FUNCTION_BLOCK UCT_PreTratamento_HMI (* Service Interface Function Block Type *)
  (* Standard: 61499-2 *)
  (* Version 1.5, 04/11/2026, Hidryco, Hidryco, 1.5: STS_LIGADO, STS_AUTOMATICO (IO List da Nereda). IHM da UCT (nomes do IThis do Pre_Tratamento antigo) *)
  PACKAGE Hidryco.HidrycoLib;
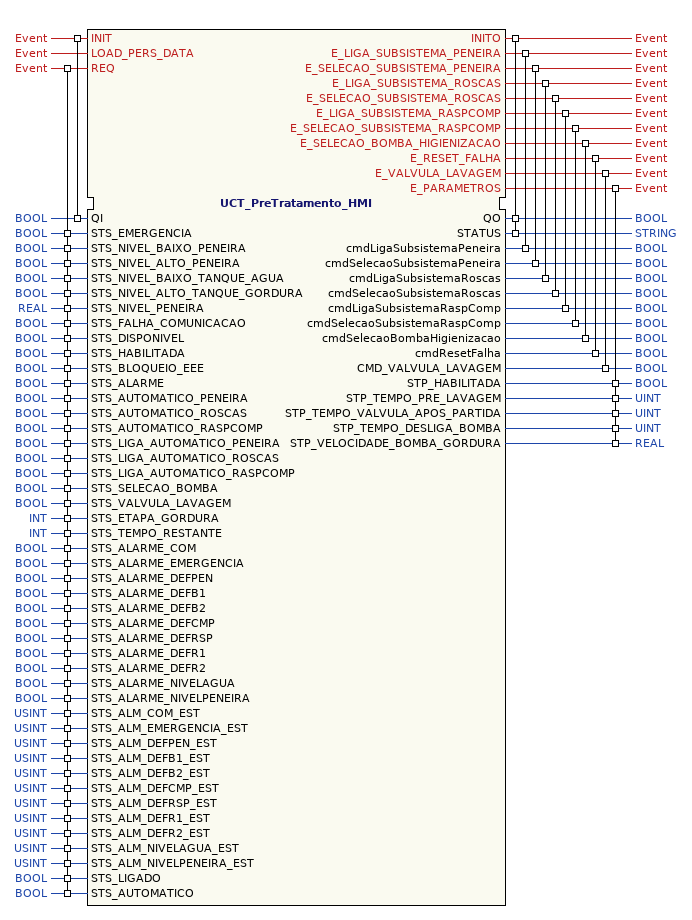
  EVENT_INPUT
    INIT WITH QI;
    LOAD_PERS_DATA; (* Reenvia os parametros persistentes *)
    REQ WITH STS_EMERGENCIA, STS_NIVEL_BAIXO_PENEIRA, STS_NIVEL_ALTO_PENEIRA, STS_NIVEL_BAIXO_TANQUE_AGUA, STS_NIVEL_ALTO_TANQUE_GORDURA, STS_NIVEL_PENEIRA, STS_FALHA_COMUNICACAO, STS_DISPONIVEL, STS_HABILITADA, STS_BLOQUEIO_EEE, STS_ALARME, STS_AUTOMATICO_PENEIRA, STS_AUTOMATICO_ROSCAS, STS_AUTOMATICO_RASPCOMP, STS_LIGA_AUTOMATICO_PENEIRA, STS_LIGA_AUTOMATICO_ROSCAS, STS_LIGA_AUTOMATICO_RASPCOMP, STS_SELECAO_BOMBA, STS_VALVULA_LAVAGEM, STS_ETAPA_GORDURA, STS_TEMPO_RESTANTE, STS_ALARME_COM, STS_ALARME_EMERGENCIA, STS_ALARME_DEFPEN, STS_ALARME_DEFB1, STS_ALARME_DEFB2, STS_ALARME_DEFCMP, STS_ALARME_DEFRSP, STS_ALARME_DEFR1, STS_ALARME_DEFR2, STS_ALARME_NIVELAGUA, STS_ALARME_NIVELPENEIRA, STS_ALM_COM_EST, STS_ALM_EMERGENCIA_EST, STS_ALM_DEFPEN_EST, STS_ALM_DEFB1_EST, STS_ALM_DEFB2_EST, STS_ALM_DEFCMP_EST, STS_ALM_DEFRSP_EST, STS_ALM_DEFR1_EST, STS_ALM_DEFR2_EST, STS_ALM_NIVELAGUA_EST, STS_ALM_NIVELPENEIRA_EST, STS_LIGADO, STS_AUTOMATICO; (* Atualizacao de status *)
  END_EVENT
  EVENT_OUTPUT
    INITO WITH QO, STATUS;
    E_LIGA_SUBSISTEMA_PENEIRA WITH cmdLigaSubsistemaPeneira;
    E_SELECAO_SUBSISTEMA_PENEIRA WITH cmdSelecaoSubsistemaPeneira;
    E_LIGA_SUBSISTEMA_ROSCAS WITH cmdLigaSubsistemaRoscas;
    E_SELECAO_SUBSISTEMA_ROSCAS WITH cmdSelecaoSubsistemaRoscas;
    E_LIGA_SUBSISTEMA_RASPCOMP WITH cmdLigaSubsistemaRaspComp;
    E_SELECAO_SUBSISTEMA_RASPCOMP WITH cmdSelecaoSubsistemaRaspComp;
    E_SELECAO_BOMBA_HIGIENIZACAO WITH cmdSelecaoBombaHigienizacao;
    E_RESET_FALHA WITH cmdResetFalha;
    E_VALVULA_LAVAGEM WITH CMD_VALVULA_LAVAGEM;
    E_PARAMETROS WITH STP_HABILITADA, STP_TEMPO_PRE_LAVAGEM, STP_TEMPO_VALVULA_APOS_PARTIDA, STP_TEMPO_DESLIGA_BOMBA, STP_VELOCIDADE_BOMBA_GORDURA;
  END_EVENT
  VAR_INPUT
    QI : BOOL;
    STS_EMERGENCIA : BOOL; (* Emergencia acionada na UCT *)
    STS_NIVEL_BAIXO_PENEIRA : BOOL; (* Nivel baixo da peneira *)
    STS_NIVEL_ALTO_PENEIRA : BOOL; (* Nivel alto da peneira *)
    STS_NIVEL_BAIXO_TANQUE_AGUA : BOOL; (* Nivel baixo do tanque de agua *)
    STS_NIVEL_ALTO_TANQUE_GORDURA : BOOL; (* Nivel alto do tanque de gordura *)
    STS_NIVEL_PENEIRA : REAL; (* Nivel da peneira (%) *)
    STS_FALHA_COMUNICACAO : BOOL; (* Falha de comunicacao com a UCT *)
    STS_DISPONIVEL : BOOL; (* UCT disponivel *)
    STS_HABILITADA : BOOL; (* UCT instalada e habilitada *)
    STS_BLOQUEIO_EEE : BOOL; (* Bloqueio do automatico da EEE Bruto (cadeia das UCTs) *)
    STS_ALARME : BOOL; (* Algum alarme da UCT *)
    STS_AUTOMATICO_PENEIRA : BOOL; (* Subsistema peneira e higienização em automatico *)
    STS_AUTOMATICO_ROSCAS : BOOL; (* Subsistema roscas em automatico *)
    STS_AUTOMATICO_RASPCOMP : BOOL; (* Subsistema raspador e compressor em automatico *)
    STS_LIGA_AUTOMATICO_PENEIRA : BOOL; (* Subsistema peneira e higienização: liga automatico em vigor *)
    STS_LIGA_AUTOMATICO_ROSCAS : BOOL; (* Subsistema roscas: liga automatico em vigor *)
    STS_LIGA_AUTOMATICO_RASPCOMP : BOOL; (* Subsistema raspador e compressor: liga automatico em vigor *)
    STS_SELECAO_BOMBA : BOOL; (* Bomba de higienizacao selecionada (FALSE bomba 1, TRUE bomba 2) *)
    STS_VALVULA_LAVAGEM : BOOL; (* Valvula de lavagem do tanque de gordura aberta *)
    STS_ETAPA_GORDURA : INT; (* Bomba de gordura: 0 parada, 1 pre-lavagem, 2 bombeando, 3 contando para desligar, 4 fora do automatico *)
    STS_TEMPO_RESTANTE : INT; (* Tempo restante (s) da etapa *)
    STS_ALARME_COM : BOOL; (* Falha de comunicação com a UCT *)
    STS_ALARME_EMERGENCIA : BOOL; (* Emergência acionada na UCT *)
    STS_ALARME_DEFPEN : BOOL; (* Defeito: Peneira rotativa *)
    STS_ALARME_DEFB1 : BOOL; (* Defeito: Bomba 1 de higienização da peneira *)
    STS_ALARME_DEFB2 : BOOL; (* Defeito: Bomba 2 de higienização da peneira *)
    STS_ALARME_DEFCMP : BOOL; (* Defeito: Compressor de ar *)
    STS_ALARME_DEFRSP : BOOL; (* Defeito: Raspador de gordura *)
    STS_ALARME_DEFR1 : BOOL; (* Defeito: Rosca 1 - horizontal *)
    STS_ALARME_DEFR2 : BOOL; (* Defeito: Rosca 2 - inclinada *)
    STS_ALARME_NIVELAGUA : BOOL; (* Nível baixo do tanque de água de higienização da UCT *)
    STS_ALARME_NIVELPENEIRA : BOOL; (* Nível alto na peneira da UCT *)
    STS_ALM_COM_EST : USINT; (* Estado do ALARM_BIT Falha de comunicação com a UCT (0 normal, 1 ativo reconhecido, 2 ativo nao reconhecido, 3 saiu nao reconhecido, 4 ativo e saiu nao reconhecido) *)
    STS_ALM_EMERGENCIA_EST : USINT; (* Estado do ALARM_BIT Emergência acionada na UCT (0 normal, 1 ativo reconhecido, 2 ativo nao reconhecido, 3 saiu nao reconhecido, 4 ativo e saiu nao reconhecido) *)
    STS_ALM_DEFPEN_EST : USINT; (* Estado do ALARM_BIT Defeito: Peneira rotativa (0 normal, 1 ativo reconhecido, 2 ativo nao reconhecido, 3 saiu nao reconhecido, 4 ativo e saiu nao reconhecido) *)
    STS_ALM_DEFB1_EST : USINT; (* Estado do ALARM_BIT Defeito: Bomba 1 de higienização da peneira (0 normal, 1 ativo reconhecido, 2 ativo nao reconhecido, 3 saiu nao reconhecido, 4 ativo e saiu nao reconhecido) *)
    STS_ALM_DEFB2_EST : USINT; (* Estado do ALARM_BIT Defeito: Bomba 2 de higienização da peneira (0 normal, 1 ativo reconhecido, 2 ativo nao reconhecido, 3 saiu nao reconhecido, 4 ativo e saiu nao reconhecido) *)
    STS_ALM_DEFCMP_EST : USINT; (* Estado do ALARM_BIT Defeito: Compressor de ar (0 normal, 1 ativo reconhecido, 2 ativo nao reconhecido, 3 saiu nao reconhecido, 4 ativo e saiu nao reconhecido) *)
    STS_ALM_DEFRSP_EST : USINT; (* Estado do ALARM_BIT Defeito: Raspador de gordura (0 normal, 1 ativo reconhecido, 2 ativo nao reconhecido, 3 saiu nao reconhecido, 4 ativo e saiu nao reconhecido) *)
    STS_ALM_DEFR1_EST : USINT; (* Estado do ALARM_BIT Defeito: Rosca 1 - horizontal (0 normal, 1 ativo reconhecido, 2 ativo nao reconhecido, 3 saiu nao reconhecido, 4 ativo e saiu nao reconhecido) *)
    STS_ALM_DEFR2_EST : USINT; (* Estado do ALARM_BIT Defeito: Rosca 2 - inclinada (0 normal, 1 ativo reconhecido, 2 ativo nao reconhecido, 3 saiu nao reconhecido, 4 ativo e saiu nao reconhecido) *)
    STS_ALM_NIVELAGUA_EST : USINT; (* Estado do ALARM_BIT Nível baixo do tanque de água de higienização da UCT (0 normal, 1 ativo reconhecido, 2 ativo nao reconhecido, 3 saiu nao reconhecido, 4 ativo e saiu nao reconhecido) *)
    STS_ALM_NIVELPENEIRA_EST : USINT; (* Estado do ALARM_BIT Nível alto na peneira da UCT (0 normal, 1 ativo reconhecido, 2 ativo nao reconhecido, 3 saiu nao reconhecido, 4 ativo e saiu nao reconhecido) *)
    STS_LIGADO : BOOL; (* UCT ligada: algum subsistema com liga-automatico (peneira, roscas ou raspador/compressor) *)
    STS_AUTOMATICO : BOOL; (* UCT em automatico: subsistema peneira em automatico *)
  END_VAR
  VAR_OUTPUT
    QO : BOOL; (* Event Output Qualifier *)
    STATUS : STRING; (* Service Status *)
    cmdLigaSubsistemaPeneira : BOOL; (* Comando cmdLigaSubsistemaPeneira *)
    cmdSelecaoSubsistemaPeneira : BOOL; (* Comando cmdSelecaoSubsistemaPeneira *)
    cmdLigaSubsistemaRoscas : BOOL; (* Comando cmdLigaSubsistemaRoscas *)
    cmdSelecaoSubsistemaRoscas : BOOL; (* Comando cmdSelecaoSubsistemaRoscas *)
    cmdLigaSubsistemaRaspComp : BOOL; (* Comando cmdLigaSubsistemaRaspComp *)
    cmdSelecaoSubsistemaRaspComp : BOOL; (* Comando cmdSelecaoSubsistemaRaspComp *)
    cmdSelecaoBombaHigienizacao : BOOL; (* Comando cmdSelecaoBombaHigienizacao *)
    cmdResetFalha : BOOL; (* Reset/reconhecimento da UCT e da bomba de gordura *)
    CMD_VALVULA_LAVAGEM : BOOL; (* Valvula de lavagem aberta (TRUE) / fechada (FALSE), so fora do automatico *)
    STP_HABILITADA : BOOL; (* UCT habilitada no bloqueio da EEE Bruto (desabilitada nao conta) *)
    STP_TEMPO_PRE_LAVAGEM : UINT; (* Tempo (s) com a valvula de lavagem aberta antes de ligar a bomba de gordura (0 = liga junto) *)
    STP_TEMPO_VALVULA_APOS_PARTIDA : UINT; (* Tempo (s) que a valvula fica aberta depois que a bomba liga (0 = fecha na partida) *)
    STP_TEMPO_DESLIGA_BOMBA : UINT; (* Tempo (s) que a bomba de gordura continua ligada depois que o nivel alto do tanque abaixa *)
    STP_VELOCIDADE_BOMBA_GORDURA : REAL; (* Velocidade da bomba de gordura em automatico (Hz) *)
  END_VAR
  SERVICE /
    SEQUENCE 
    END_SEQUENCE
  END_SERVICE
END_FUNCTION_BLOCK
